(* IEC 61131-3 sources: JingjiangArm/moonboxpro_arm_8.4/Application/Application/任务列表/CommTask, 5 files *)

(* ---- KS_CRC.st ---- *)
(*@CES
Name=KS_CRC
Type=FunctionBlock
TypeGuid=6f9dac99-8de1-4efc-8465-68ac443b7d08
Guid=c4c7953d-06dd-403a-ba97-b7ea9fcb71b0
HasDeclaration=True
HasImplementation=True
*)
{DECLARATION}
FUNCTION KS_CRC : WORD
VAR_INPUT
	i_pbyBuf: POINTER TO BYTE :=0;
	i_dwLen: DWORD;
	i_pdwSumResult: POINTER TO DWORD := 0;
END_VAR
VAR
	dwN: DWORD;
	wMask: WORD;
	wResult: WORD;
	dwSumResult: DWORD;
	pbyTemp: POINTER TO BYTE := 0;
END_VAR
{IMPLEMENTATION}

pbyTemp:= i_pbyBuf;
wResult:= 0;
dwSumResult:= 0;
FOR dwN:=1 TO i_dwLen BY 1 DO
	dwSumResult:= dwSumResult+(pbyTemp^);
	wMask:= CRC_DICTIONARY[WORD_TO_INT((wResult XOR BYTE_TO_WORD(pbyTemp^)) AND 16#FF)];
	wResult:= wMask XOR SHR(wResult,8);
	pbyTemp:= pbyTemp+1;
END_FOR
IF i_pdwSumResult<>0 THEN
	i_pdwSumResult^:= dwSumResult;
END_IF
KS_CRC:= wResult;

(* ---- KS_FillUnitMailboxCmd_DN.st ---- *)
(*@CES
Name=KS_FillUnitMailboxCmd_DN
Type=FunctionBlock
TypeGuid=6f9dac99-8de1-4efc-8465-68ac443b7d08
Guid=71378417-e57d-41a2-ab76-6caecfcdbb3a
HasDeclaration=True
HasImplementation=True
*)
{DECLARATION}
FUNCTION KS_FillUnitMailboxCmd_DN : INT
VAR_INPUT
	i_pstStParam_Mailbox: POINTER TO StParam_Mailbox;
	i_pstStUnitParam_Save: POINTER TO StUnitParam_Save;
	i_pstStUnitParam_UnSave: POINTER TO StUnitParam_UnSave;
END_VAR
VAR
	iResult: INT;
END_VAR
{IMPLEMENTATION}
iResult:= 0;
IF i_pstStParam_Mailbox<>0 AND i_pstStUnitParam_Save<>0 THEN
	i_pstStParam_Mailbox^.dwSemaphore						:= SEMA_DOWNLOAD;
	i_pstStParam_Mailbox^.dwPlateAdjustmentProf             := 0;
	i_pstStParam_Mailbox^.iRapidAdjProf_h                  	:= 0;
	i_pstStParam_Mailbox^.iGateSa                      	    := i_pstStUnitParam_Save^.iGateSa;
	i_pstStParam_Mailbox^.iGateSaEx                     	:= i_pstStUnitParam_Save^.iGateSaEx;
	i_pstStParam_Mailbox^.rAdjust_V                     	:= i_pstStUnitParam_Save^.rAdj_V;
	i_pstStParam_Mailbox^.rAdjust_H                     	:= i_pstStUnitParam_Save^.rAdj_H;
	i_pstStParam_Mailbox^.dwFlag_Ctl                    	:= i_pstStUnitParam_Save^.dwFlag_Ctl;
	i_pstStParam_Mailbox^.dwFlag_Sts                    	:= i_pstStUnitParam_Save^.dwFlag_Sts;
	i_pstStParam_Mailbox^.wButtonFun_Lamp               	:= i_pstStUnitParam_Save^.wButtonFun_Lamp;
	i_pstStParam_Mailbox^.dwSlaveBtn_HMI                	:= i_pstStUnitParam_Save^.dwSlaveBtn_HMI;
	i_pstStParam_Mailbox^.rStep_Pressure_Prn_Net        	:= i_pstStUnitParam_Save^.rStep_Pressure_Prn_Net;
	i_pstStParam_Mailbox^.rLong_Step_Roller_Pressure    	:= i_pstStUnitParam_Save^.rLong_Step_Roller_Pressure;
	i_pstStParam_Mailbox^.rShort_Step_Roller_Pressure   	:= i_pstStUnitParam_Save^.rShort_Step_Roller_Pressure;
	i_pstStParam_Mailbox^.wAirInletWindDoorValue        	:= i_pstStUnitParam_Save^.byHotBlower_AO;
	i_pstStParam_Mailbox^.wAirExhaustWindDoorValue      	:= i_pstStUnitParam_Save^.wAirExhaustWindDoorValue;
	i_pstStParam_Mailbox^.wAirReturnWindDoorValue       	:= i_pstStUnitParam_Save^.wAirReturnWindDoorValue;
	i_pstStParam_Mailbox^.dwCtlBits_UnitBaseCraft       	:= i_pstStUnitParam_Save^.dwCtlBits_UnitBaseCraft;
	i_pstStParam_Mailbox^.wHz_UnitInkRoller_ManuallySet 	:= REAL_TO_WORD(i_pstStUnitParam_Save^.rHz_UnitInkRoller_ManuallySet*100.0);
	i_pstStParam_Mailbox^.wCoeff_UnitInkRoller_Auto     	:= REAL_TO_WORD(i_pstStUnitParam_Save^.rCoeff_UnitInkRoller_Auto*100.0);
	i_pstStParam_Mailbox^.wHz_UnitScraper_ManuallySet   	:= REAL_TO_WORD(i_pstStUnitParam_Save^.rHz_UnitScraper_ManuallySet*100.0);
	i_pstStParam_Mailbox^.wCoeff_UnitScraper_Auto       	:= REAL_TO_WORD(i_pstStUnitParam_Save^.rCoeff_UnitScraper_Auto*100.0);
	i_pstStParam_Mailbox^.wHz_UnitHotWind               	:= REAL_TO_WORD(i_pstStUnitParam_Save^.rHz_UnitHotWind_ManuallySet*100.0);
	i_pstStParam_Mailbox^.wHz_UnitHotWind_2             	:= REAL_TO_WORD(i_pstStUnitParam_Save^.rHz_UnitHotWind_2_ManuallySet*100.0);
	i_pstStParam_Mailbox^.wSV_UnitTemCtl                	:= REAL_TO_WORD(i_pstStUnitParam_Save^.rSV_UnitTemCtl*100.0);
	i_pstStParam_Mailbox^.wUnit_output_I                	:= i_pstStUnitParam_UnSave^.wUnit_output_I;
	i_pstStParam_Mailbox^.wUnit_output_II               	:= i_pstStUnitParam_UnSave^.wUnit_output_II;
	//xi.hy//新增
	i_pstStParam_Mailbox^.bySignalSelect          				:= i_pstStUnitParam_Save^.bySignalSelect;
	i_pstStParam_Mailbox^.rOffset_T1          				:= i_pstStUnitParam_Save^.rOffset_T1;
	i_pstStParam_Mailbox^.rSource_Light_T1                  := i_pstStUnitParam_Save^.rSource_Light_T1;
	i_pstStParam_Mailbox^.rBias_T1          				:= i_pstStUnitParam_Save^.rBias_T1;
	i_pstStParam_Mailbox^.rBrightness_Light_T1              := i_pstStUnitParam_Save^.rBrightness_Light_T1;
	i_pstStParam_Mailbox^.rOffset_T2          				:= i_pstStUnitParam_Save^.rOffset_T2;
	i_pstStParam_Mailbox^.rSource_Light_T2                  := i_pstStUnitParam_Save^.rSource_Light_T2;
	i_pstStParam_Mailbox^.rBias_T2          				:= i_pstStUnitParam_Save^.rBias_T2;
	i_pstStParam_Mailbox^.rBrightness_Light_T2              := i_pstStUnitParam_Save^.rBrightness_Light_T2;

ELSE
	iResult:= -1;
END_IF
KS_FillUnitMailboxCmd_DN:= iResult;

(* ---- KS_FillUnitPduCmd_DN.st ---- *)
(*@CES
Name=KS_FillUnitPduCmd_DN
Type=FunctionBlock
TypeGuid=6f9dac99-8de1-4efc-8465-68ac443b7d08
Guid=77974849-7491-458e-a676-23f819d30e72
HasDeclaration=True
HasImplementation=True
*)
{DECLARATION}
FUNCTION KS_FillUnitPduCmd_DN : INT
VAR_INPUT
	i_iUnitId: INT; (* 色组id *)
	i_iGrpId_Comm: INT;(*系ID*)
	i_iCmdId: INT; (* 目前收纳61,62 *)
	i_wAxis_RollerDn: WORD;
	i_wAxis_Alarm_Prn: WORD;
	i_wComplexFlag_AxisInching: WORD;
	i_wComplexFlag_Linkage: WORD;
	i_pstStSysParam: POINTER TO StSysParam;
	i_pstStParam_PDU_Dn: POINTER TO StParam_PDU_Dn;
END_VAR
VAR
	iResult: INT;
	dwSum_Tmp: DWORD;
	pstStCMD_91: POINTER TO StPdu_Dn_91;
	pstStCMD_92: POINTER TO StPdu_Dn_92;
	pstStCMD_93: POINTER TO StPdu_Dn_93;
	pstStCMD_94: POINTER TO StPdu_Dn_94;
	pstStCMD_95: POINTER TO StPdu_Dn_95;
	pstStUnitParam_Save: POINTER TO StUnitParam_Save;
	pstStUnitParam_UnSave: POINTER TO StUnitParam_UnSave;
	uiCtl_Sample: UINT;
	iN: INT;
	iM:INT;
	byTemp: BYTE;
	dwTemp: DWORD;
	byGrpId: BYTE;
	uiTempCtl: UINT;

	dwControlComplexBits : DWORD;
	//xi.hy2026.5.9.105658
	pstStRSVUnitParam_UnSave:POINTER TO StRSV_UnitParam_UnSave;
	pstStRSVUnitParam_Save:POINTER TO StRSV_UnitParam_Save;
END_VAR
{IMPLEMENTATION}
iResult:= 0;
IF KS_IsValidUnitNR(i_iUnitId) AND(*判断轴号有效的函数*)
	(i_iGrpId_Comm=1 OR i_iGrpId_Comm=2) AND
	i_pstStSysParam<>0 AND
	i_pstStParam_PDU_Dn<>0 THEN(* 入口参数ok *)

	pstStUnitParam_Save:= ADR(i_pstStSysParam^.astStUnitParam_Save[i_iUnitId]);
	pstStUnitParam_UnSave:= ADR(i_pstStSysParam^.astStUnitParam_UnSave[i_iUnitId]);
	//xi.hy2026.5.9.102547
	pstStRSVUnitParam_UnSave:=ADR(i_pstStSysParam^.astStRSV_UnitParam_UnSave[i_iUnitId]);
	pstStRSVUnitParam_Save:=ADR(i_pstStSysParam^.astStRSV_UnitParam_Save[i_iUnitId]);
	//xi.hy
	IF pstStUnitParam_Save<>0 AND pstStUnitParam_UnSave<>0 AND pstStRSVUnitParam_UnSave<>0 AND pstStRSVUnitParam_Save<>0 THEN
		CASE i_iCmdId OF
		91:
			pstStCMD_91:= ADR(i_pstStParam_PDU_Dn^.abyPayload);
			IF pstStCMD_91<>0 THEN
				i_pstStParam_PDU_Dn^.byPkgId:= INT_TO_BYTE(i_iCmdId);

				pstStCMD_91^.byUnitId				    	:= (INT_TO_BYTE(i_iUnitId))+shl(INT_TO_byte(i_iGrpId_Comm),7);
				pstStCMD_91^.rGirth_Sam				        := pstStUnitParam_Save^.rGirth_Sam;
				pstStCMD_91^.uiNum_Sam				        := pstStUnitParam_Save^.uiNum_Sam;
				pstStCMD_91^.uiDen_Sam				        := pstStUnitParam_Save^.uiDen_Sam;
				pstStCMD_91^.byCurrUsrLevel			        := i_pstStSysParam^.stStSysParam_UnSave.byCurrUsrLevel;
				pstStCMD_91^.iCompanyId				        := i_pstStSysParam^.stStSysParam_Save.iCustomerId;
				pstStCMD_91^.byLanguageId			        := i_pstStSysParam^.stStSysParam_Save.byLanguageId;
				pstStCMD_91^.byMinutes_ScrAutoSleep	        := i_pstStSysParam^.stStSysParam_Save.byMinutes_ScrSaver;
				pstStCMD_91^.wUnit_input_I			        := pstStUnitParam_UnSave^.wUnit_input_I;
				pstStCMD_91^.wUnit_input_II                 := pstStUnitParam_UnSave^.wUnit_input_II;
				pstStCMD_91^.wUnit_input_III                := pstStUnitParam_UnSave^.wUnit_input_III;
				pstStCMD_91^.wVelocity				        := REAL_TO_WORD(i_pstStSysParam^.astStGrpParam_UnSave[i_iGrpId_Comm].rVel_Cur*10.0);
				pstStCMD_91^.wVel_Axis                      := REAL_TO_WORD(pstStUnitParam_UnSave^.rAxisVel_PrnRoller*10.0);
				pstStCMD_91^.wAxis_RollerDn                 := i_wAxis_RollerDn;
				pstStCMD_91^.wAxis_Alarm_Prn                := i_wAxis_Alarm_Prn;
				pstStCMD_91^.dwAlarmCode				    := 0;
				pstStCMD_91^.wComplexFlag_AxisInching       := i_wComplexFlag_AxisInching;
				pstStCMD_91^.wComplexFlag_Linkage      		:= i_wComplexFlag_Linkage;
				//2026.04.10.151219 修改 dwAxisFlags_Estop
				//pstStCMD_91^.wComplexFlag_Estop	       		:= 0;
				pstStCMD_91^.wComplexFlag_Estop	       		:= i_pstStSysParam^.astStRSV_GrpParam_UnSave[i_iGrpId_Comm].dwAxisFlags_Estop;
				pstStCMD_91^.wHMI_SwitchSts		          	:= 0;
				pstStCMD_91^.wSts_HorzManuPreReg	      	:= pstStUnitParam_UnSave^.wSts_HorzManuPreReg;
				pstStCMD_91^.iPos_HorzManuPreReg	    	:= pstStUnitParam_UnSave^.iPos_HorzManuPreReg;

				byGrpId:= pstStUnitParam_Save^.byGrpId;
				pstStCMD_91^.bySts_Machine.0				:= i_pstStSysParam^.astStGrpParam_UnSave[byGrpId].xFlag_Print;
				pstStCMD_91^.bySts_Machine.1			:= 0;  //设备类型 0：凹印 暂时没找到合适的判断条件 先写0
				pstStCMD_91^.byErrSts_V	:= 0;//从站暂时只用纵向状态
				pstStCMD_91^.byErrSts_V.0:= pstStUnitParam_UnSave^.xArcErrIsAlarm_V;
				pstStCMD_91^.byErrSts_V.1:= pstStUnitParam_UnSave^.xArcErrIsLost_V;
				pstStCMD_91^.byErrSts_V.2:= pstStUnitParam_UnSave^.xArcErrIsFake_V;
// 				pstStCMD_91^.byErrSts_V.4:= pstStUnitParam_UnSave^.xArcErrIsAlarm_H;
// 				pstStCMD_91^.byErrSts_V.5:= pstStUnitParam_UnSave^.xArcErrIsLost_H;
// 				pstStCMD_91^.byErrSts_V.6:= pstStUnitParam_UnSave^.xArcErrIsFake_H;
//
				//2025.11.15.132421|增加低通滤波频率下发
				pstStCMD_91^.uilowpasscutoff_hz:= pstStUnitParam_Save^.uilowpasscutoff_hz;
				i_pstStParam_PDU_Dn^.wCHK:=
					KS_CRC(
						ADR(i_pstStParam_PDU_Dn^),
						SIZEOF(i_pstStParam_PDU_Dn^)-SIZEOF(i_pstStParam_PDU_Dn^.wCHK),
						ADR(dwSum_Tmp));
			ELSE
				iResult:= -i_iCmdId;
			END_IF
		92:
			pstStCMD_92:= ADR(i_pstStParam_PDU_Dn^.abyPayload);
			IF pstStCMD_92<>0 THEN
				i_pstStParam_PDU_Dn^.byPkgId:= INT_TO_BYTE(i_iCmdId);
				pstStCMD_92^.iCurveViewMaxRange		  		:= i_pstStSysParam^.stStSysParam_Save.iCurveViewMaxRange;
				pstStCMD_92^.bySignalGain                   := pstStUnitParam_Save^.bySignalGain;
				pstStCMD_92^.byMarkTypeId                   := INT_TO_BYTE(pstStUnitParam_Save^.iMarkTypeId);
				pstStCMD_92^.byMarkArrangeModalId           := INT_TO_BYTE(pstStUnitParam_Save^.iMarkArrangeMode);
				pstStCMD_92^.byFakeThreshold_V              := pstStUnitParam_Save^.byFakeThreshold_V;
				pstStCMD_92^.byFakeThreshold_H              := pstStUnitParam_Save^.byFakeThreshold_H;
				pstStCMD_92^.rAlarm_V                       := pstStUnitParam_Save^.rAlr_V;
				pstStCMD_92^.rAlarm_H                       := pstStUnitParam_Save^.rAlr_H;
				//2026.4.11.151525 变量替换
				//pstStCMD_92^.byAve_v_extra_V                := pstStUnitParam_Save^.byAvg_V;
				pstStCMD_92^.byAve_v_extra_V                := pstStUnitParam_Save^.byAve_v_extra;
				pstStCMD_92^.byAve_v_extra_H                := pstStUnitParam_Save^.byAvg_H;
				pstStCMD_92^.iGateWidthPhy                  := pstStUnitParam_Save^.iGateWidthPhy;
				pstStCMD_92^.byTriangleMark_SideC           := i_pstStSysParam^.astStGrpParam_Save[i_iGrpId_Comm].byTriMark_SideC;
				pstStCMD_92^.byTriangleMark_SideB           := i_pstStSysParam^.astStGrpParam_Save[i_iGrpId_Comm].byTriMark_SideB;
				pstStCMD_92^.bySysSamplePrecision           := i_pstStSysParam^.astStGrpParam_Save[i_iGrpId_Comm].bySysSamplePrecision;
				pstStCMD_92^.byArcFineSampleType            := i_pstStSysParam^.astStGrpParam_Save[i_iGrpId_Comm].byArcFineSampleType;
				uiTempCtl:= 0;
				uiTempCtl.0:= TRUE;

				IF g_iMachineryType	= MACHINERYTYPE_FELXO_INLINE_ONEBOTOMROLLER THEN
					IF pstStUnitParam_UnSave^.xSamRev_BottomRoller THEN(*采样反转*)
						uiTempCtl.1:= TRUE;
					END_IF
				ELSE
					IF pstStUnitParam_UnSave^.xSamRev_PrnRoller THEN(*采样反转*)
						uiTempCtl.1:= TRUE;
					END_IF
				END_IF

				IF pstStUnitParam_Save^.uiNum_Sam= pstStUnitParam_Save^.uiDen_Sam THEN(*直驱*)
					uiTempCtl.2:= TRUE;
				END_IF
				IF pstStUnitParam_Save^.dwFlag_Ctl.9 THEN(*±10V*)
					uiTempCtl.15:= TRUE;
				END_IF
				pstStUnitParam_UnSave^.iSampleCfgParam_ctl:= UINT_TO_INT(uiTempCtl);

				pstStCMD_92^.iSampleCfgParam_ctl            := pstStUnitParam_UnSave^.iSampleCfgParam_ctl;
				pstStCMD_92^.byColorIdCurrent               := pstStUnitParam_UnSave^.byColorIdCurrent;
				pstStCMD_92^.byColorIdFollow                := pstStUnitParam_Save^.byFollowColorId;
				pstStCMD_92^.abyColorIdList[i_iUnitId]	    := 0;
				//pstStCMD_92^.bySignalSelect                 := pstStUnitParam_Save^.bySignalSelect;
				pstStCMD_92^.xEnable_Arc                    := pstStUnitParam_Save^.xEnable_arc;
				//xi.hy2026.5.9.103716
				pstStCMD_92^.wDirAndMode_FiberMove                    := SHL(BYTE_TO_WORD(pstStRSVUnitParam_UnSave^.byFiberMoveMode),8) OR pstStRSVUnitParam_UnSave^.byFiberMoveDir;
				pstStCMD_92^.uiVel_FiberMove						:=REAL_TO_UINT(pstStRSVUnitParam_UnSave^.rFiberMoveVel*10);
				pstStCMD_92^.uiDistanceOut_FiberMove						:=REAL_TO_UINT(pstStRSVUnitParam_UnSave^.rFiberMoveDistanceOut*10);
				pstStCMD_92^.uiPulsePerCycle_FiberMove						:=pstStRSVUnitParam_Save^.uiFiberMovePulsePerCycle;

				i_pstStParam_PDU_Dn^.wCHK:=
				KS_CRC(
					ADR(i_pstStParam_PDU_Dn^),
					SIZEOF(i_pstStParam_PDU_Dn^)-SIZEOF(i_pstStParam_PDU_Dn^.wCHK),
					ADR(dwSum_Tmp));
			ELSE
				iResult:= -i_iCmdId;
			END_IF

		93:
			pstStCMD_93:= ADR(i_pstStParam_PDU_Dn^.abyPayload);
			IF pstStCMD_93<>0 THEN
				i_pstStParam_PDU_Dn^.byPkgId:= INT_TO_BYTE(i_iCmdId);
//2025.11.12.132025 | 赋值错误
				//pstStCMD_93^.dwControlComplexBits	   		:= pstStUnitParam_Save^.dwCtlBits_UnitBaseCraft;
				pstStCMD_93^.dwControlComplexBits	   		:= dwControlComplexBits;
				pstStCMD_93^.wHz_UnitInkRoller_CurrWR       := REAL_TO_WORD(pstStUnitParam_UnSave^.rHz_UnitInkRoller_CurrWR*100.0);
				pstStCMD_93^.wHz_UnitScraper_CurrWR         := REAL_TO_WORD(pstStUnitParam_UnSave^.rHz_UnitScraper_CurrWR*100.0);
				pstStCMD_93^.wHz_UnitHotWind_CurrWR         := REAL_TO_WORD(pstStUnitParam_UnSave^.rHz_UnitHotWind_CurrWR*100.0);
				pstStCMD_93^.wHz_UnitHotWind2_CurrWR        := REAL_TO_WORD(pstStUnitParam_UnSave^.rHz_UnitHotWind2_CurrWR*100.0);
				pstStCMD_93^.rPV_UnitTemCtl                 := pstStUnitParam_UnSave^.rPV_UnitTemCtl;
				pstStCMD_93^.wSTS_UnitTemCtl                := pstStUnitParam_UnSave^.wSTS_UnitTemCtl;
//2026.02.07.141335增加扭矩和转速
				pstStCMD_93^.iTorque_NetRoller				:= i_pstStSysParam^.astStRSV_UnitParam_UnSave[i_iUnitId].iTorque_NetRoller;
				pstStCMD_93^.iTorque_PrnRoller				:= i_pstStSysParam^.astStRSV_UnitParam_UnSave[i_iUnitId].iTorque_PrnRoller;
				pstStCMD_93^.iTorque_BottomRoller				:= i_pstStSysParam^.astStRSV_UnitParam_UnSave[i_iUnitId].iTorque_BottomRoller;
				pstStCMD_93^.iTorque_Prn_PressRoller_M				:= i_pstStSysParam^.astStRSV_UnitParam_UnSave[i_iUnitId].iTorque_Prn_Press_M;
				pstStCMD_93^.iTorque_Prn_PressRoller_G				:= i_pstStSysParam^.astStRSV_UnitParam_UnSave[i_iUnitId].iTorque_Prn_Press_G;
				pstStCMD_93^.iTorque_Net_PressRoller_M				:= i_pstStSysParam^.astStRSV_UnitParam_UnSave[i_iUnitId].iTorque_Net_Press_M;
				pstStCMD_93^.iTorque_Net_PressRoller_G				:= i_pstStSysParam^.astStRSV_UnitParam_UnSave[i_iUnitId].iTorque_Net_Press_G;

				pstStCMD_93^.iVel_PrnRoller	:= i_pstStSysParam^.astStRSV_UnitParam_UnSave[i_iUnitId].iRpm_PrnRoller;
				pstStCMD_93^.iVel_NetRoller	:= i_pstStSysParam^.astStRSV_UnitParam_UnSave[i_iUnitId].iRpm_NetRoller;
				pstStCMD_93^.iVel_BottomRoller	:= i_pstStSysParam^.astStRSV_UnitParam_UnSave[i_iUnitId].iRpm_BottomRoller;
				//xi.hy2026.5.9.104711
				pstStCMD_93^.uiDistancePerCycle_FiberMove:=REAL_TO_UINT(pstStRSVUnitParam_Save^.rFiberMoveDistancePerCycle*100);

				i_pstStParam_PDU_Dn^.wCHK:=
				KS_CRC(
					ADR(i_pstStParam_PDU_Dn^),
					SIZEOF(i_pstStParam_PDU_Dn^)-SIZEOF(i_pstStParam_PDU_Dn^.wCHK),
					ADR(dwSum_Tmp));
			ELSE
				iResult:= -i_iCmdId;
			END_IF

		94:
			pstStCMD_94:= ADR(i_pstStParam_PDU_Dn^.abyPayload);
			IF pstStCMD_94<>0 THEN
				i_pstStParam_PDU_Dn^.byPkgId:= INT_TO_BYTE(i_iCmdId);

				pstStCMD_94^.rPos_M_Prn_HandWheelCtl		 := 0;
				pstStCMD_94^.rPos_G_Prn_HandWheelCtl         := 0;
				pstStCMD_94^.rPos_M_Net_HandWheelCtl         := 0;
				pstStCMD_94^.rPos_G_Net_HandWheelCtl         := 0;
				pstStCMD_94^.rPos_PrnRoller_Pressure_M       := pstStUnitParam_UnSave^.rPos_PrnRoller_Pressure_M;
				pstStCMD_94^.rPos_PrnRoller_Pressure_G       := pstStUnitParam_UnSave^.rPos_PrnRoller_Pressure_G;
				pstStCMD_94^.rPos_NetRoller_Pressure_M       := pstStUnitParam_UnSave^.rPos_NetRoller_Pressure_M;
				pstStCMD_94^.rPos_NetRoller_Pressure_G       := pstStUnitParam_UnSave^.rPos_NetRoller_Pressure_G;
				pstStCMD_94^.byCtlId_HandWheel               := 0;
				pstStCMD_94^.byCtlSts_HandWheel              := 0;
				pstStCMD_94^.wAxis_Alarm_Net                 := 0;
				pstStCMD_94^.wAxis_Alarm_Bottom              := 0;
				pstStCMD_94^.wAxis_Alarm_Prn_M               := 0;
				pstStCMD_94^.wAxis_Alarm_Prn_G               := 0;
				pstStCMD_94^.wAxis_Alarm_Net_M               := 0;
				pstStCMD_94^.wAxis_Alarm_Net_G               := 0;
				pstStCMD_94^.wAxis_Alarm_Other               := 0;

				i_pstStParam_PDU_Dn^.wCHK:=
				KS_CRC(
					ADR(i_pstStParam_PDU_Dn^),
					SIZEOF(i_pstStParam_PDU_Dn^)-SIZEOF(i_pstStParam_PDU_Dn^.wCHK),
					ADR(dwSum_Tmp));
			ELSE
				iResult:= -i_iCmdId;
			END_IF

		95:
			pstStCMD_95:= ADR(i_pstStParam_PDU_Dn^.abyPayload);
			IF pstStCMD_95<>0 THEN
				i_pstStParam_PDU_Dn^.byPkgId:= INT_TO_BYTE(i_iCmdId);
				(*2026.03.17.134758全自动套印*)
				pstStCMD_95^.byWidth_Mark_Max:= i_pstStSysParam^.astStRSV_UnitParam_UnSave[i_iUnitId].byWidth_Mark_Max;
				pstStCMD_95^.byWidth_Mark_Min:= i_pstStSysParam^.astStRSV_UnitParam_UnSave[i_iUnitId].byWidth_Mark_Min;
				pstStCMD_95^.byMaxGap:= i_pstStSysParam^.astStRSV_UnitParam_UnSave[i_iUnitId].byMaxGap;
				pstStCMD_95^.bySimilarityThreshold:= i_pstStSysParam^.astStRSV_UnitParam_UnSave[i_iUnitId].bySimilarityThreshold;
				pstStCMD_95^.bySpotWidth:=i_pstStSysParam^.astStRSV_UnitParam_UnSave[i_iUnitId].bySpotWidth;
				//pstStCMD_95^.bySignalType:= i_pstStSysParam^.astStRSV_UnitParam_UnSave[i_iUnitId].bySignalType;

				(*	bit0: xFlag_FindFirstMark; bit1: xFlag_FindPreMark; bit2: xFlag_AutoAdjust_Start*)
				pstStCMD_95^.byFlag_CommFromMaster:= i_pstStSysParam^.astStRSV_UnitParam_UnSave[i_iUnitId].byFlag_CommFromMaster;
				(*2026.05.20.192958||wang.xy添加内外滑窗系数通讯*)
				pstStCMD_95^.byInnerCoff:=  i_pstStSysParam^.astStRSV_UnitParam_UnSave[i_iUnitId].byInnerCoff;
				pstStCMD_95^.byOuterCoff:=  i_pstStSysParam^.astStRSV_UnitParam_UnSave[i_iUnitId].byOuterCoff;

				pstStCMD_95^.byMeanOffset:= i_pstStSysParam^.astStRSV_UnitParam_UnSave[i_iUnitId].byMeanOffset;
				FOR  iM:= 1 TO 4 BY 1 DO
					pstStCMD_95^.aiCurModeMidPoint[iM]:=i_pstStSysParam^.astStRSV_UnitParam_UnSave[i_iUnitId].aiCurModeMidPoint[iM];
					pstStCMD_95^.abyCurModeRadius[iM]:=i_pstStSysParam^.astStRSV_UnitParam_UnSave[i_iUnitId].abyCurModeRadius[iM];
					pstStCMD_95^.aiPreModeMidPoint[iM]:=i_pstStSysParam^.astStRSV_UnitParam_UnSave[i_iUnitId].aiPreModeMidPoint[iM];
					pstStCMD_95^.abyPreModeRadius[iM]:=i_pstStSysParam^.astStRSV_UnitParam_UnSave[i_iUnitId].abyPreModeRadius[iM];
				END_FOR
				//pstStCMD_95^.abyRsv_95[1] := 0;
//2026.5.7.161737增加波形美化
				pstStCMD_95^.xRsMorphFilter:= i_pstStSysParam^.astStRSV_UnitParam_Save[i_iUnitId].xRsMorphFilter;
				i_pstStParam_PDU_Dn^.wCHK:=
				KS_CRC(
					ADR(i_pstStParam_PDU_Dn^),
					SIZEOF(i_pstStParam_PDU_Dn^)-SIZEOF(i_pstStParam_PDU_Dn^.wCHK),
					ADR(dwSum_Tmp));
			ELSE
				iResult:= -i_iCmdId;
			END_IF	ELSE
			iResult:= -2;
		END_CASE
	END_IF
ELSE
	iResult:= -1;
END_IF
KS_FillUnitPduCmd_DN:= iResult;

(* ---- KS_GetNumOfDwordUsed.st ---- *)
(*@CES
Name=KS_GetNumOfDwordUsed
Type=FunctionBlock
TypeGuid=6f9dac99-8de1-4efc-8465-68ac443b7d08
Guid=eabd948f-bf57-46f0-b6b9-e9b06f242a41
HasDeclaration=True
HasImplementation=True
*)
{DECLARATION}
FUNCTION KS_GetNumOfDwordUsed : WORD
VAR_INPUT
	i_dwBytesNum				: DWORD;
END_VAR
VAR
	wResult						: WORD;
END_VAR
{IMPLEMENTATION}
wResult:= DWORD_TO_WORD(SHR(i_dwBytesNum, 2));
IF (i_dwBytesNum AND DWORD#3)<>0 THEN
	wResult:= wResult+1;
END_IF
KS_GetNumOfDwordUsed:= wResult;

(* ---- PRG_COMM.st ---- *)
(*@CES
Name=PRG_COMM
Type=FunctionBlock
TypeGuid=6f9dac99-8de1-4efc-8465-68ac443b7d08
Guid=489c5597-ab28-4682-ade4-96da00764186
HasDeclaration=True
HasImplementation=True
*)
{DECLARATION}
PROGRAM PRG_COMM
VAR
	iN:INT;(*循环变量*)
	iStationId:INT;(*通信站号*)
	stStProtocol_PDU_Up_Rd:StParam_Pdu_Up;//当前收到的实时数据PDU
	pstStCMD_F05_: POINTER TO StPdu_Up_05;
	pbyTemp:POINTER TO BYTE := 0;
	dwCheckSumVal:DWORD;
	wCHK_Up_Calc:WORD;
	diTempVal:DINT;
	tmCURR: TIME;
	tmPduSnt_LastTime: TIME; (* pdu发送的最后时间 *)
	xFlag_CmdQueueInitialized: BOOL := FALSE; (* 命令轮询初始化标志 *)
	pstStUnitCmdQueue_Tmp: POINTER TO StUnitCmdQueue; (* 命令轮询体 *)
	astStUnitCmdQueue: ARRAY [1..MAX_UNIT_NUM] OF StUnitCmdQueue := [MAX_UNIT_NUM((byCmdNum:= 0, byCmdIdx:= 1))]; (* 命令轮询结构 *)
	byIDX_Tmp: BYTE;
	byMAX_Tmp: BYTE;
	iRtn: INT;
//	iUnitNR: INT;
	abyBuf_PduCmd_snd: ARRAY [1..MAX_PDU_CMD_BYTES_DN] OF BYTE; (* 2021.12.4.154353/hdp/写入 *)
	dwDO_Tmp: DWORD; (* 数字量输出临时变量 *)
	dwOFST: DWORD;
	dwOFST2: DWORD;
	pstStUnitParam_Save: POINTER TO StUnitParam_Save;
	pstStUnitParam_UnSave: POINTER TO StUnitParam_UnSave;

	pastStParam_Mailbox: POINTER TO ARRAY [1..MAX_UNIT_NUM] OF StParam_Mailbox := 0;
	pstStParam_Mailbox_Tmp: POINTER TO StParam_Mailbox; (* 用以套用Mailbox通讯协议/2021.12.4.135959/hdp *)
	abyBuf_MailboxPkg_rcv: ARRAY [1..MAILBOX_PKG_MAX_BYTES] OF BYTE; (* Mailbox通讯的接收内存空间 *)
	axNeedUpdateParam_Malilbox: ARRAY [1..MAX_UNIT_NUM] OF BOOL:= [MAX_UNIT_NUM(0)];
	stStParam_Mailbox_Tmp: StParam_Mailbox;
	astStParam_Mailbox_snd: ARRAY [1..MAX_UNIT_NUM] OF StParam_Mailbox;
	astStParam_Mailbox_out: ARRAY [1..MAX_UNIT_NUM] OF StParam_Mailbox;
	abyBuf_MailboxPkg_snd: ARRAY [1..MAILBOX_PKG_MAX_BYTES] OF BYTE; (* Mailbox通讯的发送内存空间 *)
	pstStParam_Mailbox: POINTER TO StParam_Mailbox;
	pastStParam_Mailbox_proof: POINTER TO ARRAY [1..MAX_UNIT_NUM] OF StParam_Mailbox := 0;
	pdwSEMA: POINTER TO DWORD := 0;
	atmUnitMailboxLastSynchronized: ARRAY [1..MAX_UNIT_NUM] OF TIME := [MAX_UNIT_NUM(T#0MS)];
	diTMP: DINT;
	iUnitId_Tmp: INT;(* 色组id *)
	diValue_Tmp: DINT;(* 提交的数据 *)
	pastStProtocol_Mailbox_proof: POINTER TO ARRAY [1..MAX_UNIT_NUM] OF StParam_Mailbox := 0;
	i_xRunlogEnable: BOOL := FALSE;(* 2021.12.29.200725/hdp/增加的运行日志使能标志/不影响单次gt指令调用失败的打印信息 *)
//	i_pstStTravelLogRec: POINTER TO StTravelLogRec := 0; (* 日志入口 *)
	xSynchronized_SpecialParam: BOOL;
	udiresult : UDINT;
	iUnitId: INT;
	iGrpId: INT;
	iAxisTypeId: INT;
	axFlag_Comm_ReadEn: ARRAY [1..MAX_UNIT_NUM] OF BOOL;
	xInit_Comm_HMI: BOOL;
	abyBuf_UDP_Unit_rec: ARRAY [1..MAX_UNIT_NUM,1..MAILBOX_PKG_MAX_BYTES] OF BYTE;
	abyBuf_UDP_Unit_snd: ARRAY [1..MAX_UNIT_NUM,1..MAILBOX_PKG_MAX_BYTES] OF BYTE;
	abyBuf_UDP_Unit_rcv: ARRAY [1..MAX_UNIT_NUM,1..MAILBOX_PKG_MAX_BYTES] OF BYTE;
	abyBuf_UDP_Unit_rcv_Use_Tmp: ARRAY [1..MAILBOX_PKG_MAX_BYTES] OF BYTE;

	axFlag_DataCmd: ARRAY [1..MAX_UNIT_NUM] OF BOOL;
	abyRdDataNum: ARRAY [1..MAX_UNIT_NUM] OF BYTE;
	astStParam_UnitHMI485_Wr_81: ARRAY [1..MAX_UNIT_NUM] OF StParam_UnitHMI485_Wr_81;
	astStParam_UnitHMI485_Wr_82: ARRAY [1..MAX_UNIT_NUM] OF StParam_UnitHMI485_Wr_82;
	astStParam_UnitHMI485_Wr_83: ARRAY [1..MAX_UNIT_NUM] OF StParam_UnitHMI485_Wr_83;

	astStParam_UnitHMI485_WrRd: ARRAY [1..MAX_UNIT_NUM] OF StParam_UnitHMI485_WrRd;
	astStParam_UnitHMI485_WrRd_Rec: ARRAY [1..MAX_UNIT_NUM] OF StParam_UnitHMI485_WrRd;
	astStParam_UnitHMI485_Rd: ARRAY [1..MAX_UNIT_NUM] OF StParam_UnitHMI485_Rd;
	axFlag_Rd_OR_WrRd: ARRAY [1..MAX_UNIT_NUM] OF BOOL;
	aiStep_Comm: ARRAY [1..MAX_UNIT_NUM] OF INT;
	diTemp: DINT;
	xInit:BOOL:=FALSE;
	dwTest:DWORD;
	iRtn1: INT;
	iRtn2: INT;
	iCnt_Comm_To_gLink_II: INT;
	iCnt_Comm_To_UdpHmi: INT;
	iUnitId_To_Hmi: INT;
	xPreAcc_Ratio: BOOL;
	xPreDec_Ratio: BOOL;
	(*读取粗采样数据2025.8.14.094918*)
	iUMax_Tmp: INT;
	iUid_Tmp: INT;
	iLastId: INT;
	xReDirectedCurrUnit: BOOL;
	aiRtnCode: ARRAY [1..20] OF INT;
	iRoundSampleFlag: INT;
	pDataTest:POINTER TO BYTE;
	iM: INT;
	iGrp: INT;
	aiMarkTypeId: ARRAY [1..2] OF INT := [2(-1)]; (* A/B系标记排列选择 *)
	aiMarkArrangeId: ARRAY [1..2] OF INT := [2(-1)]; (* A/B系标记排列 *)
	lrTempVal: LREAL;
	pstStGrpParam_Save: POINTER TO StGrpParam_Save;
	pstStGrpParam_UnSave: POINTER TO StGrpParam_UnSave;
	wAxis_RollerDn				:WORD  ;(*轴压辊状态(bit0-1U,bit15-16U)*)
	wAxis_Alarm_Prn				:WORD  ;(*色组版辊报警状态(bit0-1U,bit15-16U)*)
	dwAlarmCode					:DWORD ;(*轴报警码*)
	wComplexFlag_AxisInching	:WORD  ;(*所有轴的单运行状态*)
	wComplexFlag_Linkage		:WORD  ;(*所有轴的联动状态*)
	wComplexFlag_Estop			:DWORD ;(*所有轴的急停状态*)
	byGrpId: BYTE;
	axSynchronizedFlag			: ARRAY [1..MAX_UNIT_NUM] OF BOOL:= [MAX_UNIT_NUM(FALSE)];
	abyHorzManu_HMI_Pre			: ARRAY [1..MAX_UNIT_NUM] OF BYTE;
	adwCtlBits_UnitBaseCraft_Temp	: ARRAY [1..MAX_UNIT_NUM] OF DWORD;

	aiCntInch : ARRAY [1..MAX_UNIT_NUM] OF INT;

	(*月光宝盒、月光宝盒pr设置标志@2025.8.7.220536+*)
	axRemoteSetDne				: ARRAY [1..MAX_STATION_NUM] OF  BOOL;
	axRemotSetFailed			: ARRAY [1..MAX_STATION_NUM] OF BOOL;

	adwMotorEncoder : ARRAY [1..MAX_UNIT_NUM] OF DWORD := [MAX_UNIT_NUM(4194304)];

	auiAllowMotorRpm_Max : ARRAY [1..MAX_UNIT_NUM] OF UINT := [MAX_UNIT_NUM(5000)];

//2026.1.4.175023增加子影人机通讯内容2026.1.4.175033
	iGrpIdTmp: INT;

	pdata1: POINTER TO BYTE;
	pdata2: POINTER TO BYTE;
	iK: INT;
	iLength: INT;
	xFlag_MasterChange: BOOL;
	aiCntPress : ARRAY [1..MAX_UNIT_NUM] OF INT;
	aiCntUnPress : ARRAY [1..MAX_UNIT_NUM] OF INT;
aiTime: ARRAY [1..max_unit_num] OF INT;
aiTime1: ARRAY [1..max_unit_num] OF INT;
	udiAddrRd:UDINT;

			//xi.hy
	pstStRSVUnitParam_UnSave:POINTER TO StRSV_UnitParam_UnSave;
	pstStRSVUnitParam_Save:POINTER TO StRSV_UnitParam_Save;
	xTest:BOOL;
	awState_FiberMove_bak:ARRAY [1..MAX_UNIT_NUM] OF WORD;
	fbKS_FB_ExportRSFifo2File: KS_FB_ExportRSFifo2File;(*2026.03.23.162629||wang.xy*)

	(*2026.5.7.183226lhy+*)
	dwNetTime_Act:ARRAY [1..MAX_STATION_NUM] OF DWORD;

	//2026.08.06.203155
	aiCntStop: ARRAY [1..MAX_UNIT_NUM] OF INT;
END_VAR

{IMPLEMENTATION}
IF g_iRunStepId=RUNSTEP_NormalWork AND g_dwTensionRunNum>=5 THEN
	;
ELSE
	RETURN;
END_IF
iCnt_Comm_To_gLink_II:= iCnt_Comm_To_gLink_II+1;
iCnt_Comm_To_UdpHmi:= iCnt_Comm_To_UdpHmi+1;
(*金刚通讯5ms执行周期*)
Action_Udp_Diamonds();

IF g_stStSysParam.stStSysParam_Save.dwEquipmentProf.3 THEN
(*凹印的套色用值就用版辊吧2025.9.12.163315*)

	FOR iN:= 1 TO MAX_UNIT_NUM BY 1 DO
		g_stStSysParam.astStUnitParam_Save[iN].rGirth_Sam := g_stStSysParam.astStUnitParam_Save[iN].rGirth_PrnRoller;
		g_stStSysParam.astStUnitParam_Save[iN].uiNum_Sam := g_stStSysParam.astStUnitParam_Save[iN].uiNum_PrnRoller;
		g_stStSysParam.astStUnitParam_Save[iN].uiDen_Sam := g_stStSysParam.astStUnitParam_Save[iN].uiDen_PrnRoller;
	END_FOR

	IF iCnt_Comm_To_gLink_II>= 3 THEN
		iCnt_Comm_To_gLink_II:= 0;
Action_gLink_II_Input();

		Action_GLINKII_COMM();
Action_gLink_II_Output();

		Action_RdSampleData();//S2025.08.23.200014+

	END_IF
	iCnt_Comm_To_UdpHmi:= 0;
ELSIF g_stStSysParam.stStSysParam_Save.dwEquipmentProf.2 OR g_stStSysParam.stStSysParam_Save.dwEquipmentProf.5 THEN

	//2025.12.24.162857 | + | bai.zy | 秦华的采样周长比较特殊
	IF g_stStSysParam.stStSysParam_Save.iCustomerId = CUSTOMERNAME_QINHUA THEN
		FOR iN:= 1 TO MAX_UNIT_NUM BY 1 DO
			g_stStSysParam.astStUnitParam_Save[iN].rGirth_Sam := g_stStSysParam.astStUnitParam_Save[iN].rGirth_PrnRoller;
			g_stStSysParam.astStUnitParam_Save[iN].uiNum_Sam := REAL_TO_UINT(UINT_TO_REAL(g_stStSysParam.astStUnitParam_Save[iN].uiNum_BottomRoller) * g_stStSysParam.astStUnitParam_Save[iN].rGirth_PrnRoller *1000/
								g_stStSysParam.astStGrpParam_Save[1].rGirth_BottomRoller);(* 减速比-电机端 *);//g_stStSysParam.astStUnitParam_Save[iN].uiNum_PrnRoller;
			g_stStSysParam.astStUnitParam_Save[iN].uiDen_Sam := 1000;//g_stStSysParam.astStUnitParam_Save[iN].uiDen_PrnRoller;
		END_FOR
	ELSE
		//2025.12.01.164356 | +
		FOR iN:= 1 TO MAX_UNIT_NUM BY 1 DO
			g_stStSysParam.astStUnitParam_Save[iN].rGirth_Sam := g_stStSysParam.astStUnitParam_Save[iN].rGirth_PrnRoller;
			g_stStSysParam.astStUnitParam_Save[iN].uiNum_Sam := g_stStSysParam.astStUnitParam_Save[iN].uiNum_PrnRoller;
			g_stStSysParam.astStUnitParam_Save[iN].uiDen_Sam := g_stStSysParam.astStUnitParam_Save[iN].uiDen_PrnRoller;
		END_FOR
	END_IF

	IF iCnt_Comm_To_gLink_II>= 3 THEN
		iCnt_Comm_To_gLink_II:= 0;
Action_gLink_II_Input();

		Action_GLINKII_COMM();
Action_gLink_II_Output();

		Action_RdSampleData();//S2025.08.23.200014+

	END_IF

	IF iCnt_Comm_To_UdpHmi>= 2 THEN
		//Action_Udp_UnitHMI();
		iCnt_Comm_To_UdpHmi:= 0;
	END_IF
	//iCnt_Comm_To_gLink_II:= 0;
END_IF
Action_SyncParamToSample();

(*2026.5.14.091424屏蔽了
//2025.12.16.154650 | 异站编码器新增加的功能测试，目前先放在这里，暂时还没有库，等待中。。。。。。
FOR iN:=1 TO g_stStSysParam.stStSysParam_Save.iUnitMaxNum BY 1 DO
	pstStUnitParam_Save:=ADR(g_stStSysParam.astStUnitParam_Save[iN]);
	IF 	pstStUnitParam_Save^.iStationId<>-1 THEN(*存在控制站号*)
//2026.03.11.093012 | + | 同步获取编码器位数和最大转速的功能 下面的这一段改成自动的，不使用强制了，已经在秦华验证过
		IF NOT axRemoteSetDne[iN] THEN
			//2026.02.23.161037 | + | 通过flash获取编码器位数
			udiAddrRd:= 289;(* Nos *)
			iRtn :=GTN_RN_GetFlashParamInfo(
					cardIndex:= 1,
					station_id:= pstStUnitParam_Save^.iStationId,
					axis:= 1,
					addr:= udiAddrRd,
					pData:= ADR(adwMotorEncoder[iN]));
			(*目前只支持这两种编码器@2025.12.5.151451*)
			IF adwMotorEncoder[iN]<>4194304 AND
				adwMotorEncoder[iN]<>16777216 THEN
				adwMotorEncoder[iN]:=4194304;
			END_IF

			//2026.02.23.161037 | + | 通过flash获取最高转速
			udiAddrRd:= 80;(* Nos *)
			iRtn :=GTN_RN_GetFlashParamInfo(
					cardIndex:= 1,
					station_id:= pstStUnitParam_Save^.iStationId,
					axis:= 1,
					addr:= udiAddrRd,
					pData:= ADR(auiAllowMotorRpm_Max[iN]));
		END_IF
		KS_SetRemoteEncParam(FALSE,(*使用异站编码器@true 使用本地编码器*)
						g_abyStationList_CommKSCR[iN],//pstStUnitParam_Save^.iStationId,
						adwMotorEncoder[iN],
						auiAllowMotorRpm_Max[iN],//REAL_TO_UINT(pstStAxisParam^.rAllowMotorRpm_Max),
						DINT_TO_DWORD(gc_diVirEncPPR_New),(*有可能根据套色采样精度修改*)
						ADR(axRemoteSetDne[iN]),
						ADR(axRemotSetFailed[iN]));

	ELSE
		axRemoteSetDne[iN]:=FALSE;
		axRemotSetFailed[iN]:=FALSE;
	END_IF
END_FOR
*)
